//---------------------------------------------------------------------------------------------------------------
//
//  HAUD 2026.11.07
//
//  - fb_TicketConductor
//  -----------------------------
//  - detects new entry in the linked list
//    - forwards the received entry to cyclic linked list
//    - cyclic linked list is then sending the ticket abroad.
//
//  - Ctrl / State for you to use (uses instance ctrl/state pair)
//    - this is simply a ENABLE / DISABLE class
//    - the input list is simply checked for (count > 0)
//  - this conductor has no transport process
//  - this conductor is used for sending tickets to cyclic list strucutres
//---------------------------------------------------------------------------------------------------------------
FUNCTION_BLOCK fb_TicketConductor
VAR
  _nConductor             : E_INSTANCE := E_INSTANCE.INSTANCE_CONDUCTOR; // msg device identifier, in case you instantiate more than one conductor
  _stCtrl                 : REFERENCE TO ST_INSTANCE_CTRL;
  _stState                : REFERENCE TO ST_INSTANCE_STATE;

  _eCmd,
  _eCmdOld                : E_INSTANCE_CMD;       // commands for local state machine
  _eStateInstance         : E_INSTANCE_STATE;     // local state machine for infeed procedure

  _eResult                : E_PROGRESS;           // result for methods
  _eStateProgress         : E_PROGRESS;           // substate for local state machine

  _eInit                  : E_PROGRESS;           // startup
  _eCheck                 : E_INSTANCE_CHECK;     // pointer checks

  // the outbox
  _stListCtrl             : REFERENCE TO ST_LIST_CTRL;
  _stListState            : REFERENCE TO ST_LIST_STATE;
  _stListDataInput        : REFERENCE TO ST_LIST_NODE_DATA;

  // the inbox
  _ItfTicketList          : I_Process_LinkedList;
  _ResultTicketList       : ST_PROCESS_LIST_RESULT;   // internal list results
  _DeleteResult           : ST_PROCESS_LIST_RESULT;   // last job executed

  _stMsg                  : ST_Message;
  _MessageLevel           : E_MessageType := E_MessageType.eMessageInfo;
END_VAR

//-----------------------------------------------------------------------------
//-----------------------------------------------------------------------------
// check pointer and interface
// set message device identification
//-----------------------------------------------------------------------------
IF NOT Check() THEN 
  RETURN; 
END_IF
//-----------------------------------------------------------------------------
// check command
//-----------------------------------------------------------------------------
_eCmd                                         := _stCtrl.Cmd;
IF (_eCmd <> _eCmdOld)
THEN
  CASE _eCmd
  OF
    E_INSTANCE_CMD.INIT:
      _eStateInstance                         := E_INSTANCE_STATE.NULL;
      _eStateProgress                         := E_PROGRESS.PROGRESS_INIT;
  END_CASE
  CmdLog();
  _eCmdOld                                    := _eCmd;
END_IF
//-----------------------------------------------------------------------------
//-----------------------------------------------------------------------------
// state machine for ProcessConductor work
//-----------------------------------------------------------------------------
CASE _eStateInstance
OF
  E_INSTANCE_STATE.NULL:
    // first cycle startup
    _eInit                                    := E_PROGRESS.PROGRESS_INVALID;
    _eStateProgress                           := E_PROGRESS.PROGRESS_INIT;
    _eStateInstance                           := E_INSTANCE_STATE.INIT;


  E_INSTANCE_STATE.INIT:
    //-------------------------------------------------------------------------
    CASE _eStateProgress
    OF
    // E_INSTANCE_STATE.INIT:
    //-------------------------------------------------------------------------
      E_PROGRESS.PROGRESS_INIT:
        IF (_ItfTicketList <> 0)
        THEN
          _eStateProgress                     := E_PROGRESS.PROGRESS_BUSY;
        END_IF
    // E_INSTANCE_STATE.INIT:
    //-------------------------------------------------------------------------
      E_PROGRESS.PROGRESS_BUSY:
        IF _ItfTicketList.InitList()
        THEN
          IF (_stListState.Init <> E_PROGRESS.PROGRESS_DONE)
          THEN
            _stListCtrl.Cmd                   := E_LIST_CTRL.LIST_CTRL_NULL;
            _eStateProgress                   := E_PROGRESS.PROGRESS_PREPARE;
          ELSE
            _eInit                            := E_PROGRESS.PROGRESS_DONE;
  
            _eStateInstance                   := E_INSTANCE_STATE.DISABLED;
            _eStateProgress                   := E_PROGRESS.PROGRESS_BUSY;
          END_IF
        ELSE
          _eStateProgress                     := E_PROGRESS.PROGRESS_ERROR;
        END_IF
    // E_INSTANCE_STATE.INIT:
    //-------------------------------------------------------------------------
      E_PROGRESS.PROGRESS_PREPARE:
        _stListCtrl.Cmd                       := E_LIST_CTRL.LIST_CTRL_INIT;

        IF (_stListState.Init = E_PROGRESS.PROGRESS_DONE)
        THEN
          _stListCtrl.Cmd                     := E_LIST_CTRL.LIST_CTRL_NULL;
          _eStateInstance                     := E_INSTANCE_STATE.DISABLED;
          _eStateProgress                     := E_PROGRESS.PROGRESS_BUSY;
          _eInit                              := E_PROGRESS.PROGRESS_DONE;

        ELSIF (_stListState.Init = E_PROGRESS.PROGRESS_ERROR)
        THEN
          _eStateProgress                     := E_PROGRESS.PROGRESS_ERROR;
        END_IF
    END_CASE
END_CASE
//-----------------------------------------------------------------------------
// DISABLED:
//  - clear local list result data
//  - wait for enable from the outside
//-----------------------------------------------------------------------------
CASE _eStateInstance
OF
  E_INSTANCE_STATE.DISABLED:
    //-------------------------------------------------------------------------
    CASE _eStateProgress
    OF
      E_PROGRESS.PROGRESS_BUSY:
        CASE _eCmd
        OF
          E_INSTANCE_CMD.ENABLE:              // turn it on!!
            _stListCtrl.Cmd                   := E_LIST_CTRL.LIST_CTRL_NULL;

            _eStateInstance                   := E_INSTANCE_STATE.DETECTION;
            _eStateProgress                   := E_PROGRESS.PROGRESS_BUSY;
  
            IF (_MessageLevel > E_MessageType.eMessageInfo)
            THEN
              _stMsg.eType                    := E_MessageType.eMessageVerbose;
              _stMsg.eSubdevice               := e_Subdevice.Instance_ProcessConductor;
              _stMsg.iErrorNumber             := 0;
              _stMsg.sText                    := concat(TO_STRING(_eStateInstance), ': ');
              _stMsg.sText                    := concat(_stMsg.sText, TO_STRING(_eStateProgress));
              f_MessageSet(_stMsg);
            END_IF
        END_CASE
    END_CASE
END_CASE
//-----------------------------------------------------------------------------
// DETECTION: 
//  - check inked list and GetHead()
//  - copy job data
//  - switch on process
//-----------------------------------------------------------------------------
CASE _eStateInstance
OF
  E_INSTANCE_STATE.DETECTION:
    //-------------------------------------------------------------------------
    CASE _eStateProgress
    OF
      E_PROGRESS.PROGRESS_BUSY:
        IF (_eCmd = E_INSTANCE_CMD.DISABLE)
        THEN
          _eStateInstance                     := E_INSTANCE_STATE.DISABLED;
          _eStateProgress                     := E_PROGRESS.PROGRESS_BUSY;
  
        ELSIF (_ItfTicketList.Count > 0)
        THEN
          // get new job order for my process
          // the list results carries information about who and where
          _ResultTicketList                   := _ItfTicketList.GetHead();
  
          IF (_ResultTicketList.wState <> 0)
          THEN
            // error in list results must not appear
            // if you land here, there is somethng wrong with the initialization or configuration of the linked list
            _eStateProgress                   := E_PROGRESS.PROGRESS_ERROR;
  
            _stMsg.eType                      := E_MessageType.eMessageError;
            _stMsg.eSubdevice                 := e_Subdevice.Instance_ProcessConductor;
            _stMsg.iErrorNumber               := _ResultTicketList.wState;
            _stMsg.sText                      := concat(TO_STRING(_eStateInstance), ': _ResultTicketList.wState: ');
            _stMsg.sText                      := concat(_stMsg.sText, TO_STRING(_eStateProgress));
            f_MessageSet(_stMsg);
  
          ELSE
            IF (_MessageLevel > E_MessageType.eMessageError)
            THEN
              _stMsg.eType                    := E_MessageType.eMessageInfo;
              _stMsg.eSubdevice               := e_Subdevice.Instance_ProcessConductor;
              _stMsg.iErrorNumber             := _ResultTicketList.stData.wTarget;
              _stMsg.sText                    := concat(TO_STRING(_eStateInstance), ': ');
              _stMsg.sText                    := concat(_stMsg.sText, '_ResultTicketList.stData.wTarget: ');
              _stMsg.sText                    := concat(_stMsg.sText, BitsToString(_ResultTicketList.stData.wTarget));
              f_MessageSet(_stMsg);
            END_IF
  
            IF (_ResultTicketList.stData.wTarget > 0)
            THEN
              _eStateProgress                 := E_PROGRESS.PROGRESS_PREPARE;
  
              IF (_MessageLevel > E_MessageType.eMessageEmpty)
              THEN
                _stMsg.eType                  := E_MessageType.eMessageBatch;
                _stMsg.eSubdevice             := e_Subdevice.Instance_ProcessConductor;
                _stMsg.iErrorNumber           := 0;
                _stMsg.sText                  := concat(TO_STRING(_eStateProgress), ': ');
                _stMsg.sText                  := concat(_stMsg.sText, TO_STRING(e_message_batch.MSG_BATCH_JOB_STARTED));
                f_MessageSet(_stMsg);
              END_IF
            ELSE
              _ResultTicketList               := _ItfTicketList.RemoveHeadValue();

              IF (_ResultTicketList.wState <> 0)
              THEN
                _stMsg.eType                  := E_MessageType.eMessageError;
                _stMsg.eSubdevice             := e_Subdevice.Instance_ProcessConductor;
                _stMsg.iErrorNumber           := _ResultTicketList.wState;
                _stMsg.sText                  := concat(TO_STRING(_eStateProgress), ': _ResultTicketList.wState: ');
                _stMsg.sText                  := concat(_stMsg.sText, BitsToString(_ResultTicketList.wState));
                f_MessageSet(_stMsg);

                _eStateProgress               := E_PROGRESS.PROGRESS_ERROR;
              END_IF
            END_IF
  
            // check target mask for entries
            IF NOT (_ResultTicketList.stData.wTarget > 0)
            THEN
              _stMsg.eType                    := E_MessageType.eMessageWarning;
              _stMsg.eSubdevice               := e_Subdevice.Process_LinkedList_CheckData;
              _stMsg.iErrorNumber             := 666;
              _stMsg.sText                    := concat(TO_STRING(_eStateInstance), ': ');
              _stMsg.sText                    := concat(_stMsg.sText, '_ResultTicketList.stData.wTarget: ');
              _stMsg.sText                    := concat(_stMsg.sText, BitsToString(_ResultTicketList.stData.wTarget));
              f_MessageSet(_stMsg);
            END_IF
          END_IF
        END_IF

      E_PROGRESS.PROGRESS_PREPARE:
        // check process target plausibility
        IF NOT (_ResultTicketList.stData.nProcessId > 0) OR
           NOT (_ResultTicketList.stData.nProcessId < E_INSTANCE.INSTANCE_MAX)
        THEN
          _ResultTicketList                   := _ItfTicketList.RemoveHeadValue();
  
          IF (_ResultTicketList.wState <> 0)
          THEN
            _stMsg.eType                      := E_MessageType.eMessageError;
            _stMsg.eSubdevice                 := e_Subdevice.Instance_ProcessConductor;
            _stMsg.iErrorNumber               := _ResultTicketList.wState;
            _stMsg.sText                      := concat(TO_STRING(_eStateProgress), ': _ResultTicketList.wState: ');
            _stMsg.sText                      := concat(_stMsg.sText, BitsToString(_ResultTicketList.wState));
            f_MessageSet(_stMsg);

            _eStateProgress                   := E_PROGRESS.PROGRESS_ERROR;
          END_IF

          _stMsg.eType                        := E_MessageType.eMessageError;
          _stMsg.eSubdevice                   := e_Subdevice.Process_LinkedList_CheckData;
          _stMsg.iErrorNumber                 := 6666;
          _stMsg.sText                        := concat(TO_STRING(_eStateInstance), ': ');
          _stMsg.sText                        := concat(_stMsg.sText, '_ResultTicketList.stData.nProcessId: ');
          _stMsg.sText                        := concat(_stMsg.sText, TO_STRING(_ResultTicketList.stData.nProcessId));
          f_MessageSet(_stMsg);
  
        ELSE
          IF (_MessageLevel > E_MessageType.eMessageInfo)
          THEN
            _stMsg.eType                      := E_MessageType.eMessageVerbose;
            _stMsg.eSubdevice                 := e_Subdevice.Instance_ProcessConductor;
            _stMsg.iErrorNumber               := _ResultTicketList.stData.nProcessId;
            _stMsg.sText                      := concat(TO_STRING(_eStateInstance), ': _ResultTicketList.stData.nProcessId: ');
            _stMsg.sText                      := concat(_stMsg.sText, TO_STRING(_ResultTicketList.stData.nProcessId));
            f_MessageSet(_stMsg);
          END_IF

          _stListDataInput.ProcessData        := _ResultTicketList.stData;
          _DeleteResult                       := _ItfTicketList.RemoveHeadValue();
  
          IF (_DeleteResult.wState = 0)
          THEN
            _eStateInstance                   := E_INSTANCE_STATE.WORKING;
            _eStateProgress                   := E_PROGRESS.PROGRESS_BUSY;
          ELSE
            _stMsg.eType                      := E_MessageType.eMessageError;
            _stMsg.eSubdevice                 := e_Subdevice.Instance_ProcessConductor;
            _stMsg.iErrorNumber               := _DeleteResult.wState;
            _stMsg.sText                      := concat(TO_STRING(_eStateProgress), ': _DeleteResult.wState: ');
            _stMsg.sText                      := concat(_stMsg.sText, BitsToString(_DeleteResult.wState));
            f_MessageSet(_stMsg);

            _eStateProgress                   := E_PROGRESS.PROGRESS_ERROR;
          END_IF
        END_IF
    END_CASE
END_CASE
//-----------------------------------------------------------------------------
// WORKING
//  - Add ticket in target list
//  - check and log
//  - transition to finish
//-----------------------------------------------------------------------------
CASE _eStateInstance
OF
  E_INSTANCE_STATE.WORKING:
    //-------------------------------------------------------------------------
    CASE _eStateProgress
    OF
      E_PROGRESS.PROGRESS_BUSY:
        _stListCtrl.Cmd                       := E_LIST_CTRL.LIST_CTRL_ADD_TAIL;

        IF (_stListState.State = E_LIST_STATE.LIST_STATE_ADD_TAIL + E_PROGRESS.PROGRESS_DONE)
        THEN
          _stListCtrl.Cmd                     := E_LIST_CTRL.LIST_CTRL_NULL;
          _eStateInstance                     := E_INSTANCE_STATE.FINISH;
          _eStateProgress                     := E_PROGRESS.PROGRESS_BUSY;

        ELSIF (_stListState.State = E_LIST_STATE.LIST_STATE_ADD_TAIL + E_PROGRESS.PROGRESS_ERROR)
        THEN
          _eStateProgress                     := E_PROGRESS.PROGRESS_ERROR;
        END_IF
    END_CASE
END_CASE
//-----------------------------------------------------------------------------
// FINISH:
//-----------------------------------------------------------------------------
CASE _eStateInstance
OF
  E_INSTANCE_STATE.FINISH:
    //-------------------------------------------------------------------------
    CASE _eStateProgress
    OF
      E_PROGRESS.PROGRESS_BUSY:
        _eStateProgress                       := E_PROGRESS.PROGRESS_DONE;
    END_CASE
    // E_INSTANCE_STATE.FINISH:
    //-------------------------------------------------------------------------
    CASE _eStateProgress
    OF
      E_PROGRESS.PROGRESS_DONE:
        _eStateInstance                       := E_INSTANCE_STATE.DISABLED;
        _eStateProgress                       := E_PROGRESS.PROGRESS_BUSY;
    END_CASE
END_CASE
//-----------------------------------------------------------------------------
//-----------------------------------------------------------------------------
_stState.ProcessIdentity                      := _nConductor;
_stState.ProcessState                         := _eStateInstance;
_stState.ProcessProgress                      := _eStateProgress;
_stState.QueueProcessCount                    := TO_UINT(_ItfTicketList.Count);
//-----------------------------------------------------------------------------
//-----------------------------------------------------------------------------

METHOD PUBLIC BitGet : BOOL
VAR_INPUT
  inVal   : T_PROCESS;
  bitNo   : DINT;
END_VAR
VAR
  wConst : T_PROCESS := 1;
END_VAR
IF ( inVal AND SHL( wConst,TO_SINT(bitNo) MOD TO_INT(SIZEOF(T_PROCESS)*8) ) ) > 0
THEN
  BitGet := TRUE;
ELSE
  BitGet := FALSE;
END_IF
END_METHOD

METHOD BitsToString : STRING(SIZEOF(T_PROCESS)*8) // T_PROCESS to string
VAR_INPUT
  inVal       : T_PROCESS;
END_VAR
VAR
  _nx         : DINT;
  _str        : STRING(SIZEOF(T_PROCESS)*8);
END_VAR
FOR _nx := ((SIZEOF(inVal)*8)) TO 1 BY(-1)
DO
  IF (BitGet(inVal, _nx-1))
  THEN
    _str     := concat(_str, '1');
  ELSE
    _str     := concat(_str, '0');
  END_IF
END_FOR

BitsToString := _str;
END_METHOD

METHOD Check  : BOOL // call this method in the extending/inheriting class
VAR_INST
  _idx        : UINT;
END_VAR
//-----------------------------------------------------------------------------
//-----------------------------------------------------------------------------
// pointer checks
//-----------------------------------------------------------------------------
IF NOT __ISVALIDREF(_stCtrl)
THEN
  _eCheck                 := E_INSTANCE_CHECK.INVALID_INSTANCE_CONTROL_REFERENCE;
  RETURN;
END_IF

IF NOT __ISVALIDREF(_stState)
THEN
  _eCheck                 := E_INSTANCE_CHECK.INVALID_INSTANCE_STATE_REFERENCE;
  RETURN;
END_IF

IF NOT __ISVALIDREF(_stListCtrl)
THEN
  _eCheck                 := E_INSTANCE_CHECK.CTRL_CYCLIC_LIST_REFERENCE_INVALID;
  RETURN;
END_IF

IF NOT __ISVALIDREF(_stListState)
THEN
  _eCheck                 := E_INSTANCE_CHECK.STATE_CYCLIC_LIST_REFERENCE_INVALID;
  RETURN;
END_IF

IF NOT __ISVALIDREF(_stListDataInput)
THEN
  _eCheck                 := E_INSTANCE_CHECK.DATA_CYCLIC_LIST_REFERENCE_INVALID;
  RETURN;
END_IF

IF NOT (_ItfTicketList <> 0)
THEN
  _eCheck                 := E_INSTANCE_CHECK.TICKET_LIST_ITF_INVALID;
  RETURN;
END_IF

//-----------------------------------------------------------------------------
//-----------------------------------------------------------------------------
// set message device
//-----------------------------------------------------------------------------
_stMsg.eDevice            := e_Device.Conductor + TO_UINT(_nConductor);
//-----------------------------------------------------------------------------
//-----------------------------------------------------------------------------
_eCheck                   := E_INSTANCE_CHECK.CHECK_DONE;
Check                     := TRUE;
END_METHOD

METHOD CmdLog

IF (_MessageLevel > E_MessageType.eMessageError)
THEN
  _stMsg.eSubdevice       := e_Subdevice.Instance_ProcessConductor;
  _stMsg.iErrorNumber     := 0;
  _stMsg.sText            := concat('E_INSTANCE_CMD', '.');
  _stMsg.sText            := concat(_stMsg.sText, TO_STRING(_eCmd));
  f_MessageSet(_stMsg);
END_IF
END_METHOD

PROPERTY Ctrl : REFERENCE TO ST_INSTANCE_CTRL
SET
_stCtrl ref= Ctrl;
END_SET
END_PROPERTY

PROPERTY CyclicListCtrl : REFERENCE TO ST_LIST_CTRL
SET
_stListCtrl ref= CyclicListCtrl;
END_SET
END_PROPERTY

PROPERTY CyclicListData : REFERENCE TO ST_LIST_NODE_DATA
SET
_stListDataInput ref= CyclicListData;
END_SET
END_PROPERTY

PROPERTY CyclicListState : REFERENCE TO ST_LIST_STATE
SET
_stListState ref= CyclicListState;
END_SET
END_PROPERTY

PROPERTY MessageLevel : e_MessageType
GET
MessageLevel := _MessageLevel;
END_GET
SET
_MessageLevel := MessageLevel;
END_SET
END_PROPERTY

PROPERTY State : REFERENCE TO ST_INSTANCE_STATE
SET
_stState ref= State;
END_SET
END_PROPERTY

PROPERTY TicketLinkedList : I_Process_LinkedList
SET
_ItfTicketList := TicketLinkedList;
END_SET
END_PROPERTY

END_FUNCTION_BLOCK

(* stored: Version 1.1.0.1
   POU fb_TicketConductor: Id {b2975459-610b-4622-ae2f-021df5bebfac}, SpecialFunc None
   Method BitGet: Id {c2d83cf2-dbce-411d-a81b-1737586284e7}
   Method BitsToString: Id {f72cba2b-f8e8-4a05-bc02-5475239bcff5}
   Method Check: Id {cb3f11a1-f1a7-4ee3-af44-3681fdcfcb4b}
   Method CmdLog: Id {3965707d-6687-42ea-8ffe-d947bf5ebb46}
   Property Ctrl: Id {8d31c008-953c-4cdb-a8c4-26723f8f0e0f}
   Set Set: Id {a892d71d-b682-4094-8364-be7d9e8ec86b}
   Property CyclicListCtrl: Id {71be235e-4c27-4f6b-a895-003158074062}
   Set Set: Id {00c0aa77-d61e-46bd-b8e0-3c7cdf765c44}
   Property CyclicListData: Id {9b975f5f-3816-4b09-a847-b7fe55c01647}
   Set Set: Id {12baa5fa-1ba5-4230-a01d-c5d033de624b}
   Property CyclicListState: Id {0f63748a-bd58-40ca-8c4c-510773bc5e48}
   Set Set: Id {11e69477-81e3-4a5a-84fc-e67caf9f716b}
   Property MessageLevel: Id {c3a2d482-eeba-4134-b03b-197f0d97cb34}
   Get Get: Id {7ba8c18c-6749-4fa2-8211-ea77d590f394}
   Set Set: Id {d39bd273-7573-4d9a-afb7-0895896e2af3}
   Property State: Id {ef65cd4b-e98c-4206-888b-dafd5e0fe13a}
   Set Set: Id {3fe56f4c-ad87-4410-9959-ddf819640b22}
   Property TicketLinkedList: Id {c3042300-b508-4f79-9b52-b4795f611b89}
   Set Set: Id {4bbcf1b1-0fac-4d0a-b322-a8efa117641b} *)
